        MoveL Target_6940,v300,z10,ToolLab1AlexaReyes\WObj:=Workobject_1;
        MoveL Target_6950,v300,z10,ToolLab1AlexaReyes\WObj:=Workobject_1;
    ENDPROC
    PROC Path_210()
        MoveL Target_6960,v300,z10,ToolLab1AlexaReyes\WObj:=Workobject_1;
        MoveL Target_6970,v300,z10,ToolLab1AlexaReyes\WObj:=Workobject_1;
        MoveL Target_6980,v300,z10,ToolLab1AlexaReyes\WObj:=Workobject_1;
        MoveL Target_6990,v300,z10,ToolLab1AlexaReyes\WObj:=Workobject_1;
    ENDPROC
    PROC Path_220()
        MoveJ Target_Mant,v300,z10,ToolLab1AlexaReyes\WObj:=wobj0;
    ENDPROC
    PROC Path_230()
        MoveJ Target_7000,v100,z10,ToolLab1AlexaReyes\WObj:=Workobject_1;
        MoveJ Target_7010,v100,z10,ToolLab1AlexaReyes\WObj:=Workobject_1;
        MoveJ Target_7020,v100,z10,ToolLab1AlexaReyes\WObj:=Workobject_1;
        MoveJ Target_7030,v100,z10,ToolLab1AlexaReyes\WObj:=Workobject_1;
        MoveJ Target_7040,v100,z10,ToolLab1AlexaReyes\WObj:=Workobject_1;
    ENDPROC

ENDMODULE

--- Controller Data/IRB140_6_81/SYSPAR/EIO.cfg ---
EIO:CFG_1.0:6:1::
#
EIO_SIGNAL:

      -Name "DI_01" -SignalType "DI"

      -Name "DI_02" -SignalType "DI"

      -Name "DI_03" -SignalType "DI"

      -Name "DO_01" -SignalType "DO"

      -Name "DO_02" -SignalType "DO"

      -Name "DO_03" -SignalType "DO"

      -Name "FWD_Conveyor" -SignalType "DO"

      -Name "BWD_Conveyor" -SignalType "DO"
